FUNCTION_BLOCK ActuatorRouter IMPLEMENTS I_Actuator, I_Cyclic
VAR
    _Name   : STRING(32);
    _Source : E_DeviceSource;
    _Chosen : I_Actuator;
END_VAR
(*
    ActuatorRouter

    One I_Actuator in front of up to four candidates, chosen once by the
    site setting. Only the chosen candidate is run. A source with no
    candidate (0) is never at either end, and reports a fault.
*)

METHOD FB_init : BOOL
VAR_INPUT
    bInitRetains    : BOOL;
    bInCopyCode     : BOOL;
    Name            : STRING(32);
    Source          : E_DeviceSource;
    FinalHardware   : I_Actuator;
    SimilarHardware : I_Actuator;
    Simulation      : I_Actuator;
    Test            : I_Actuator;
END_VAR
_Name := Name;
_Source := Source;
CASE Source OF
    E_DeviceSource.FinalHardware:   _Chosen := FinalHardware;
    E_DeviceSource.SimilarHardware: _Chosen := SimilarHardware;
    E_DeviceSource.Simulation:      _Chosen := Simulation;
    E_DeviceSource.Test:            _Chosen := Test;
END_CASE
END_METHOD

METHOD PUBLIC CyclicLogic
VAR
    Cyclic : I_Cyclic;
END_VAR
IF _Chosen <> 0 AND_THEN __QUERYINTERFACE(_Chosen, Cyclic) THEN
    Cyclic.CyclicLogic();              // only the chosen candidate runs
END_IF
END_METHOD

METHOD PUBLIC Extend
IF _Chosen <> 0 THEN
    _Chosen.Extend();
END_IF
END_METHOD

METHOD PUBLIC Retract
IF _Chosen <> 0 THEN
    _Chosen.Retract();
END_IF
END_METHOD

METHOD PUBLIC Reset
IF _Chosen <> 0 THEN
    _Chosen.Reset();
END_IF
END_METHOD

PROPERTY PUBLIC IsExtended : BOOL
GET
IsExtended := _Chosen <> 0 AND_THEN _Chosen.IsExtended;
END_GET
END_PROPERTY

PROPERTY PUBLIC IsRetracted : BOOL
GET
IsRetracted := _Chosen <> 0 AND_THEN _Chosen.IsRetracted;
END_GET
END_PROPERTY

PROPERTY PUBLIC Name : STRING
GET
Name := _Name;
END_GET
END_PROPERTY

PROPERTY PUBLIC HasFault : BOOL
GET
HasFault := _Chosen = 0 OR_ELSE _Chosen.HasFault;
END_GET
END_PROPERTY

PROPERTY PUBLIC FaultText : STRING
GET
IF _Chosen = 0 THEN
    FaultText := 'No device for this source';
ELSE
    FaultText := _Chosen.FaultText;
END_IF
END_GET
END_PROPERTY

PROPERTY PUBLIC Source : E_DeviceSource
GET
Source := _Source;
END_GET
END_PROPERTY

END_FUNCTION_BLOCK

(* stored: Version 1.1.0.1, ProductVersion 3.1.4026.0
   POU ActuatorRouter: Id {0343c712-987f-45d8-8c5c-9d8f2265f44d}, SpecialFunc None
   Folder I_Actuator: Id {1c504744-3918-4f8c-9c1b-2c459a847c6b}
   Folder I_Diagnosable: Id {359cfdb6-0727-46bf-9786-6b12983feee0}
   Folder I_Resettable: Id {b9dd2623-dd13-4837-ad7a-80d781276af5}
   Folder I_Cyclic: Id {323133cf-d7c3-49bb-a612-3140ef99fd02}
   Method FB_init: Id {c39ea1b0-0146-4a58-afb3-209e0b84986f}
   Method CyclicLogic: Id {f27eb673-441e-4ea6-ac3f-9a21474d38c8}
   Method Extend: Id {4c2d5a61-bacc-4f52-b49c-8ec0ade09c92}
   Method Retract: Id {4922259b-c985-4d68-b4b5-0d83a812704d}
   Method Reset: Id {503bad84-cf40-4688-b146-1b89786dada8}
   Property IsExtended: Id {94314995-0958-453e-b7fc-9048003e645d}
   Get Get: Id {9ea89229-4cc7-4b22-8f2e-52f088b81688}
   Property IsRetracted: Id {1454d7d5-3b79-40ac-aed2-62dcec4427e1}
   Get Get: Id {bc159ccf-21b6-4f87-9eb9-518f2cca352f}
   Property Name: Id {cd8a049f-ef93-4d5d-b0ce-543a925fdfca}
   Get Get: Id {e3eca068-b5d4-4b08-9e6e-200bdee96101}
   Property HasFault: Id {ab4b31e7-5ddb-4e01-97fe-f85ed68fdab0}
   Get Get: Id {a6bc8458-7bad-425f-be3f-f6b951b7e703}
   Property FaultText: Id {15916a38-e01f-4743-b773-f1aa902a00ce}
   Get Get: Id {44767648-3c6e-4fce-8a28-b26f52260f44}
   Property Source: Id {e2a9b67b-ed78-42eb-ab87-6076fa6f6cf9}
   Get Get: Id {7cdec107-1185-46dc-ae8c-053f971be645} *)
